// TIA Portal V21 export
// export: Created 2000-01-01T00:00:00.0000000Z, ExportSetting None
FUNCTION "MCP_B6_LadFc" : Void   // FC9602, LAD
TITLE = 条件与定时
{ S7_Optimized_Access := 'TRUE' }
// stored: SetENOAutomatically false
   VAR_TEMP   // added for the SCL form of the ladder/FBD networks
      _w1 : Bool;
      _w2 : Bool;
   END_VAR
BEGIN

REGION Network 1
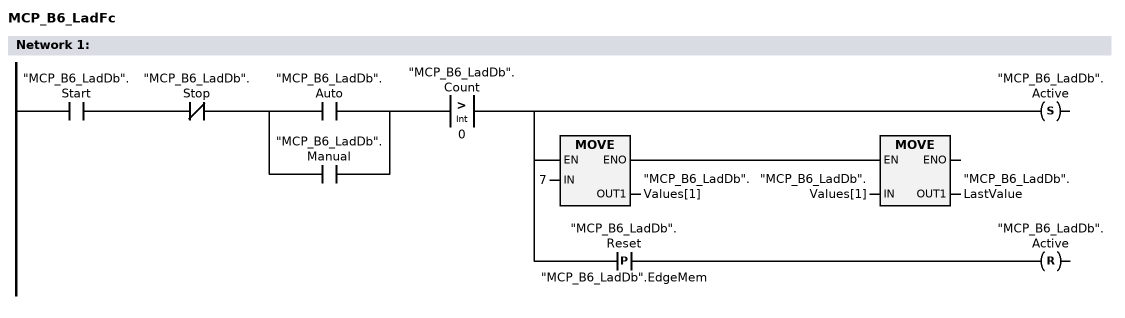
   // ENO of a box is taken as its EN; it also drops when the box reports an error
   #_w1 := "MCP_B6_LadDb".Start AND NOT "MCP_B6_LadDb".Stop AND ("MCP_B6_LadDb".Auto OR "MCP_B6_LadDb".Manual) AND ("MCP_B6_LadDb".Count > 0);
   IF #_w1 THEN
       "MCP_B6_LadDb".Active := TRUE;
       "MCP_B6_LadDb".Values[1] := 7;
       "MCP_B6_LadDb".LastValue := "MCP_B6_LadDb".Values[1];
   END_IF;
   #_w2 := "MCP_B6_LadDb".Reset AND NOT "MCP_B6_LadDb".EdgeMem;   // rising edge of "MCP_B6_LadDb".Reset
   "MCP_B6_LadDb".EdgeMem := "MCP_B6_LadDb".Reset;
   IF #_w2 THEN "MCP_B6_LadDb".Active := FALSE; END_IF;
END_REGION
END_FUNCTION
